(* PLC project v0.5.4_.project, CODESYS CODESYS V3.5 SP19 Patch 1 *)
(* stored: creationDateTime 2026-08-04T04:55:17.9088614, modificationDateTime 2026-08-04T04:54:49.1401172 *)

PROGRAM PRG_06_Outputs_LD
  VAR_OUTPUT
    PowerKeepAlive_A_RQ : BOOL;
    PowerKeepAlive_B_RQ : BOOL;
    EmergencyArming_RQ : BOOL;
    EmergencyArmingPulseActive : BOOL;
    EmergencyArmingLockoutActive : BOOL;
    ArmingSeqStep : INT;
    RedundancyTestFailed : BOOL;
    EmergencyArmingFailed : BOOL;
  END_VAR
  VAR
    M1RelayFwd : BOOL;
    instM1RelayFwd : FB_Output;
    instSafetyEmergencyManagement : FB_Safety_EmergencyManagement;
    PowerCutOffReq : BOOL;
  END_VAR

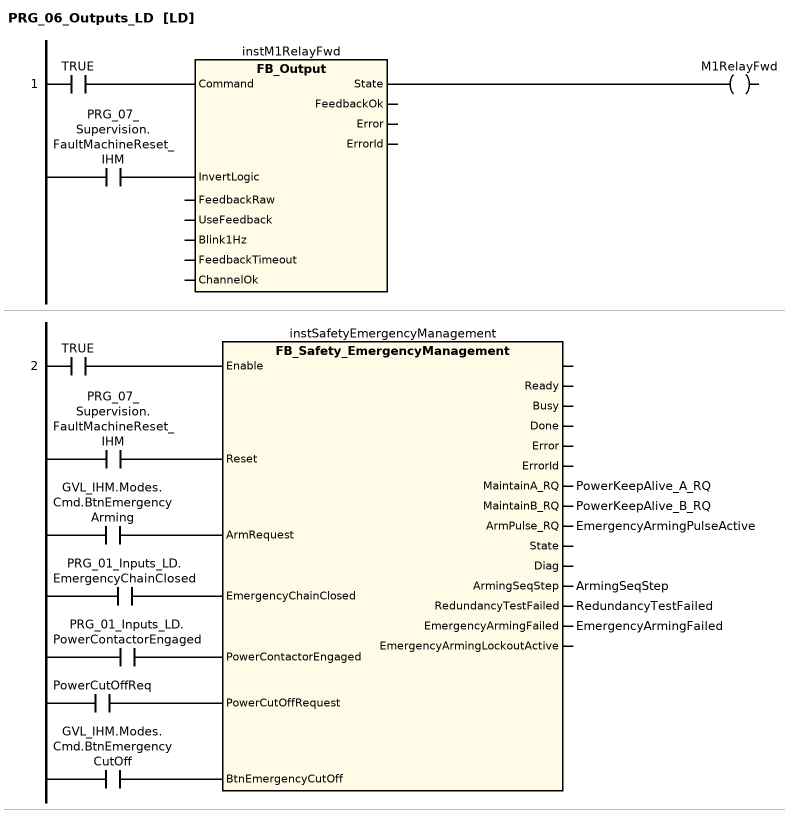
(* LD diagram, written out as Structured Text *)

instM1RelayFwd(Command := TRUE, InvertLogic := PRG_07_Supervision.FaultMachineReset_IHM, FeedbackRaw := , UseFeedback := , Blink1Hz := , FeedbackTimeout := , ChannelOk := );
M1RelayFwd := instM1RelayFwd.State;

instSafetyEmergencyManagement(Enable := TRUE, Reset := PRG_07_Supervision.FaultMachineReset_IHM, ArmRequest := GVL_IHM.Modes.Cmd.BtnEmergencyArming, EmergencyChainClosed := PRG_01_Inputs_LD.EmergencyChainClosed, PowerContactorEngaged := PRG_01_Inputs_LD.PowerContactorEngaged, PowerCutOffRequest := PowerCutOffReq, BtnEmergencyCutOff := GVL_IHM.Modes.Cmd.BtnEmergencyCutOff, MaintainA_RQ => PowerKeepAlive_A_RQ, MaintainB_RQ => PowerKeepAlive_B_RQ, ArmPulse_RQ => EmergencyArmingPulseActive, ArmingSeqStep => ArmingSeqStep, RedundancyTestFailed => RedundancyTestFailed, EmergencyArmingFailed => EmergencyArmingFailed);
END_PROGRAM
